(*
SPDX-FileCopyrightText: © 2026 Oleksandr Tiutyk <trofimich@gmail.com>
SPDX-License-Identifier: MIT
License: https://opensource.org/license/mit
*)

(*!
<summary>Orders LINT values described by generic descriptors.</summary>
<description>
Non-null addresses must reference live LINT storage. TypeClass and Size are not validated and no numeric
conversion is performed. Two null addresses compare equal; one null address sorts before a non-null address.
Descriptors are passed by value; payload remains borrowed and is not modified, cloned, released or retained.
IsMemoryOwner does not affect comparison.
</description>
*)

FUNCTION_BLOCK LIntComparer EXTENDS TOF_Core.Object IMPLEMENTS TOF_Core.IComparer
VAR_STAT
	//! <summary>Class name shared by all instances of this function block.</summary>
	{attribute 'hide'} 
	_ClassName : STRING := __POUNAME();
END_VAR

{attribute 'monitoring' := 'call'}
PROPERTY ClassName : REFERENCE TO STRING
GET
ClassName REF= _ClassName;
END_GET
END_PROPERTY

(*!
<summary>Compares the first operand with the second using this ordering strategy.</summary>
<description>
Non-null addresses must reference live LINT storage. TypeClass and Size are not validated and no numeric
conversion is performed. Two null addresses compare equal; one null address sorts before a non-null address.
Descriptors are passed by value; payload remains borrowed and is not modified, cloned, released or retained.
IsMemoryOwner does not affect comparison. Descendants cannot replace this standard ordering; implement
IComparer separately for a different ordering strategy.
</description>
*)
//!<param name="first">First descriptor; referenced storage is borrowed for the call.</param>
//!<param name="second">Second descriptor; referenced storage is borrowed for the call.</param>
{attribute "object_name" := "Compare"}
METHOD FINAL Compare : TOF_Core.COMPARISON_RESULT
VAR_INPUT
	first : TOF_Core.GENERIC_VALUE;
	second : TOF_Core.GENERIC_VALUE;
END_VAR
VAR
	leftPointer : POINTER TO LINT; 
	rightPointer : POINTER TO LINT; 
END_VAR
IF first.Address = 0 AND_THEN second.Address = 0 THEN
	Compare := TOF_Core.COMPARISON_RESULT.FIRST_EQUAL_TO_SECOND;
	RETURN;
END_IF

IF first.Address = 0 THEN
	Compare := TOF_Core.COMPARISON_RESULT.FIRST_LESS_THAN_SECOND;
	RETURN;	
END_IF

IF second.Address = 0 THEN
	Compare := TOF_Core.COMPARISON_RESULT.FIRST_GREATER_THAN_SECOND;
	RETURN;	
END_IF

leftPointer := first.Address;
rightPointer := second.Address;

IF leftPointer^ < rightPointer^ THEN
	Compare := TOF_Core.COMPARISON_RESULT.FIRST_LESS_THAN_SECOND;
ELSIF leftPointer^ > rightPointer^ THEN
	Compare := TOF_Core.COMPARISON_RESULT.FIRST_GREATER_THAN_SECOND;
ELSE
	Compare := TOF_Core.COMPARISON_RESULT.FIRST_EQUAL_TO_SECOND;	
END_IF
END_METHOD

{attribute 'monitoring' := 'call'}
PROPERTY NamespaceName : REFERENCE TO STRING
GET
NamespaceName REF= CurrentNamespace.Name;
END_GET
END_PROPERTY

{attribute 'monitoring' := 'call'}
PROPERTY SelfSize : ULINT
GET
SelfSize := XSIZEOF(THIS^);
END_GET
END_PROPERTY

END_FUNCTION_BLOCK

(* stored: Version 1.1.0.1
   POU LIntComparer: Id {6802d232-eb84-4fc6-9db7-da1a848885bb}, SpecialFunc None
   Property ClassName: Id {11696811-cbc8-4330-9b9c-34480612a1fd}
   Get Get: Id {9443910c-a564-4f25-a954-0af25c296bce}
   Method Compare: Id {16519cb2-8b2a-4d05-af51-ba14c0acf190}
   Property NamespaceName: Id {08b866a6-e0c1-4fc7-9eca-ea0da6a53d8a}
   Get Get: Id {8bc84db1-d75e-4bbf-af7b-e6873dc30080}
   Property SelfSize: Id {c25e4d6f-9f0f-4471-9ede-a23224e4040d}
   Get Get: Id {00ea876a-2583-4961-990c-bcb33b2f9770} *)
